// TIA Portal V17 export
// export: Created 2026-11-08T05:50:31.9466979Z, ExportSetting WithDefaults, DisplayName Totally Integrated Automation Portal, DisplayVersion V17, DisplayName TIA Portal Openness, DisplayVersion V17, DisplayName TIA Portal Version Control Interface, DisplayVersion V17, DisplayName STEP 7 Professional, DisplayVersion V17, DisplayName STEP 7 Safety, DisplayVersion V17, DisplayName WinCC Professional, DisplayVersion V17
TextList "Estilos"  ListRange=Decimal
  TextListEntry   EntryType=SingleValue, From=1, To=1, Text="BANDERAS"
  TextListEntry   EntryType=SingleValue, From=2, To=2, Text="MOORE"
  TextListEntry   EntryType=SingleValue, From=3, To=3, Text="MEALY"
